// TwinCAT 3 PLC project HeartbeatWatchdogTests
// ProgramVersion: 3.1.4026.22
// libraries:
//   Tc2_Standard, * (Beckhoff Automation GmbH)
//   Tc2_System, * (Beckhoff Automation GmbH)
// project tree:
//   StateMachineControl/POUs/ FB_HeartbeatWatchdog.TcPOU
//   StateMachineControl/tests/POUs/ PRG_HeartbeatWatchdogTests.TcPOU
//   StateMachineControl/tests/ TestTask.TcTTO
// (motion and I/O tree: see PLC project experimentsequencertests)
// real-time tasks:
//   TASK DriveStateTestTask: cycle T#10ms, priority 1, ADS port 350
//   TASK TestTask: cycle T#10ms, priority 2, ADS port 351

CONFIGURATION HeartbeatWatchdogTests
    RESOURCE PLC ON TwinCAT3
        TASK TestTask(INTERVAL := T#10ms, PRIORITY := 2);
        PROGRAM PRG_HeartbeatWatchdogTests WITH TestTask : PRG_HeartbeatWatchdogTests;
    END_RESOURCE
END_CONFIGURATION

// ---- StateMachineControl/tests/POUs/PRG_HeartbeatWatchdogTests.TcPOU
PROGRAM PRG_HeartbeatWatchdogTests
VAR
    watchdog : FB_HeartbeatWatchdog;
    testsExecuted : BOOL := FALSE;
    testsPassed : BOOL := FALSE;
    failureCount : UDINT := 0;
END_VAR

IF NOT testsExecuted THEN
    (* Disabled state synchronizes the counter and stays inactive. *)
    watchdog(enable := FALSE, heartbeatCounter := 10, timeoutTicks := 3);
    IF watchdog.timeout OR watchdog.tripEdge THEN
        failureCount := failureCount + 1;
    END_IF

    (* Timeout occurs on the Nth enabled call, not before it. *)
    watchdog(enable := TRUE, heartbeatCounter := 10, timeoutTicks := 3);
    IF watchdog.timeout OR watchdog.tripEdge THEN
        failureCount := failureCount + 1;
    END_IF
    watchdog(enable := TRUE, heartbeatCounter := 10, timeoutTicks := 3);
    IF watchdog.timeout OR watchdog.tripEdge THEN
        failureCount := failureCount + 1;
    END_IF
    watchdog(enable := TRUE, heartbeatCounter := 10, timeoutTicks := 3);
    IF NOT watchdog.timeout OR NOT watchdog.tripEdge THEN
        failureCount := failureCount + 1;
    END_IF

    (* A sustained timeout emits only one trip edge. *)
    watchdog(enable := TRUE, heartbeatCounter := 10, timeoutTicks := 3);
    IF NOT watchdog.timeout OR watchdog.tripEdge THEN
        failureCount := failureCount + 1;
    END_IF

    (* A heartbeat change clears timeout and rearms edge detection. *)
    watchdog(enable := TRUE, heartbeatCounter := 11, timeoutTicks := 3);
    IF watchdog.timeout OR watchdog.tripEdge THEN
        failureCount := failureCount + 1;
    END_IF
    watchdog(enable := TRUE, heartbeatCounter := 11, timeoutTicks := 3);
    watchdog(enable := TRUE, heartbeatCounter := 11, timeoutTicks := 3);
    watchdog(enable := TRUE, heartbeatCounter := 11, timeoutTicks := 3);
    IF NOT watchdog.timeout OR NOT watchdog.tripEdge THEN
        failureCount := failureCount + 1;
    END_IF

    (* Disable clears the latch; the same heartbeat can trip again after rearm. *)
    watchdog(enable := FALSE, heartbeatCounter := 11, timeoutTicks := 3);
    IF watchdog.timeout OR watchdog.tripEdge THEN
        failureCount := failureCount + 1;
    END_IF
    watchdog(enable := TRUE, heartbeatCounter := 11, timeoutTicks := 3);
    watchdog(enable := TRUE, heartbeatCounter := 11, timeoutTicks := 3);
    watchdog(enable := TRUE, heartbeatCounter := 11, timeoutTicks := 3);
    IF NOT watchdog.timeout OR NOT watchdog.tripEdge THEN
        failureCount := failureCount + 1;
    END_IF

    (* A zero timeout trips immediately when enabled. *)
    watchdog(enable := FALSE, heartbeatCounter := 20, timeoutTicks := 0);
    watchdog(enable := TRUE, heartbeatCounter := 20, timeoutTicks := 0);
    IF NOT watchdog.timeout OR NOT watchdog.tripEdge THEN
        failureCount := failureCount + 1;
    END_IF

    testsExecuted := TRUE;
    testsPassed := (failureCount = 0);
END_IF

END_PROGRAM

// ---- StateMachineControl/POUs/FB_HeartbeatWatchdog.TcPOU
FUNCTION_BLOCK FB_HeartbeatWatchdog
VAR_INPUT
    enable : BOOL;
    heartbeatCounter : UDINT;
    timeoutTicks : UDINT;
END_VAR
VAR_OUTPUT
    timeout : BOOL := FALSE;
    tripEdge : BOOL := FALSE;
END_VAR
VAR
    counterPrev : UDINT := 0;
    silenceTicks : UDINT := 0;
    tripLatched : BOOL := FALSE;
    heartbeatChanged : BOOL := FALSE;
END_VAR

tripEdge := FALSE;
heartbeatChanged := (heartbeatCounter <> counterPrev);

IF NOT enable THEN
    counterPrev := heartbeatCounter;
    silenceTicks := 0;
    tripLatched := FALSE;
ELSIF heartbeatChanged THEN
    counterPrev := heartbeatCounter;
    silenceTicks := 0;
    tripLatched := FALSE;
ELSE
    IF silenceTicks < timeoutTicks THEN
        silenceTicks := silenceTicks + 1;
    END_IF
END_IF

timeout := enable AND (silenceTicks >= timeoutTicks);
IF timeout AND NOT tripLatched THEN
    tripEdge := TRUE;
    tripLatched := TRUE;
END_IF

END_FUNCTION_BLOCK
